// TIA Portal V21 export
// export: Created 2026-11-11T00:48:08.6250651Z, ExportSetting WithDefaults, DisplayName Totally Integrated Automation Portal, DisplayVersion V21 Update 3, DisplayName STEP 7 Professional, DisplayVersion V21 Update 3, DisplayName STEP 7 Safety, DisplayVersion V21, DisplayName Tech WebApplication, DisplayVersion V21, DisplayName WinCC Basic/Comfort/Advanced, DisplayVersion V21 Update 3, DisplayName WinCC Unified, DisplayVersion V21 Update 3
FUNCTION_BLOCK "FB_Scl_sl009"   // FB37, SCL
{ S7_Optimized_Access := 'TRUE' }
VERSION : 0.1
// stored: AutoNumber true, IsIECCheckEnabled false, IsRetainMemResEnabled false, MemoryReserve 100, SetENOAutomatically false, UDAEnableTagReadback false
   VAR_INPUT
      v_t_no : Timer;
      v_s : Bool;
      v_tv : S5Time;
      v_r : Bool;
   END_VAR
   VAR_OUTPUT
      v_q : Bool;
      v_bi : Word;
   END_VAR
BEGIN
   #v_bi := S_PULSE(T_NO := #v_t_no, S := #v_s, TV := #v_tv, R := #v_r, Q => #v_q);
END_FUNCTION_BLOCK
